FUNCTION_BLOCK TcoSequencerNonAutoRestorableTest EXTENDS TcoCore._internals_TcoContext
VAR
	_callMyPlcInstance	:	BOOL := FALSE;
	_sequencer : _TcoSequencer(THIS^, eRestoreMode.None);
	_runPLCinstanceOnce : BOOL := FALSE;
	_runPLCinstanceCyclicaly : BOOL := FALSE;
	_stepID : INT := 32764;
	_enabled : BOOL;
	_stepDescription : STRING := 'Last step sequence message';	
	_runOneStep : BOOL;
	_runAllSteps : BOOL;
	_finishStep : BOOL;
	_restore : BOOL;
	_cycleCount : INT;
	_restoreCycleCount : INT;
	_init: BOOL;
END_VAR

IF _callMyPlcInstance THEN
	IF NOT _init THEN
		ContextOpen();	
		ContextClose();	
		_init := THIS^._rtc.IsValid;
	END_IF
	
	IF _restore THEN
		ContextOpen();	
		THIS^._sequencer.Restore();	
		_restoreCycleCount := _restoreCycleCount + 1;
		_restore := FALSE;
		ContextClose();	
		RETURN;
	END_IF
	
	IF _runPLCinstanceOnce AND NOT _runPLCinstanceCyclicaly THEN
		ContextOpen();	
		THIS^.PLCinstanceRun(_stepID , _enabled, _stepDescription);
		_cycleCount := _cycleCount + 1;
		_runPLCinstanceOnce := FALSE;
		ContextClose();	
	END_IF
	
	IF _runPLCinstanceCyclicaly AND NOT _runPLCinstanceOnce THEN
		ContextOpen();	
		THIS^.PLCinstanceRun(_stepID , _enabled, _stepDescription);
		_cycleCount := _cycleCount + 1;
		ContextClose();	
	END_IF
END_IF;

{attribute 'TcRpcEnable'}
METHOD ChildHasAutoRestoreEnabled : BOOL;
ChildHasAutoRestoreEnabled := _sequencer.ChildHasAutoRestoreEnabled();
END_METHOD

{attribute 'TcRpcEnable'}
METHOD ChildIsAutoRestorable : BOOL;
ChildIsAutoRestorable := _sequencer.ChildIsAutoRestorable();
END_METHOD

{attribute 'TcRpcEnable'}
METHOD CleanupPointers
_sequencer.CleanupPointers();
END_METHOD

{attribute 'TcRpcEnable'}
METHOD ClearNumberOfSteps
_sequencer.ClearNumberOfSteps();
END_METHOD

{attribute 'TcRpcEnable'}
METHOD PROTECTED ContextClose
SUPER^._Close();
END_METHOD

{attribute 'TcRpcEnable'}
METHOD ContextOpen
SUPER^._Open();
END_METHOD

{attribute 'TcRpcEnable'}
METHOD GetChildState : INT
GetChildState := _sequencer.GetChildState();
END_METHOD

{attribute 'TcRpcEnable'}
METHOD GetCurrentStepOrder : UINT
GetCurrentStepOrder := _sequencer._currentStep.Order;
END_METHOD

{attribute 'TcRpcEnable'}
METHOD GetNumberOfStepsInSequence : UINT
GetNumberOfStepsInSequence := _sequencer._numberOfStepsInSequence;
END_METHOD

{attribute 'TcRpcEnable'}
METHOD GetOrderOfTheCurrentlyEvaluatedStep : UINT
GetOrderOfTheCurrentlyEvaluatedStep := _sequencer._theOrderOfTheCurrentlyEvaluatedStep;
END_METHOD

{attribute 'TcRpcEnable'}
METHOD GetOrderOfTheCurrentlyExecutedStep : UINT
GetOrderOfTheCurrentlyExecutedStep := _sequencer._theOrderOfTheCurrentlyExecutedStep;
END_METHOD

{attribute 'TcRpcEnable'}
METHOD GetPreviousNumberOfStepsInSequence : UINT
GetPreviousNumberOfStepsInSequence := _sequencer._previousNumberOfStepsInSequence;
END_METHOD

{attribute 'TcRpcEnable'}
METHOD GetRequestStepCycle : UINT
GetRequestStepCycle := _sequencer.RequestStepCycle;
END_METHOD

{attribute 'TcRpcEnable'}
METHOD GetSequencerErrorId : INT
GetSequencerErrorId := _sequencer.GetSequencerErrorId();
END_METHOD

{attribute 'TcRpcEnable'}
METHOD GetTextOfTheMostImportantMessage : STRING(254)
GetTextOfTheMostImportantMessage := THIS^._sequencer.GetTextOfTheMostImportantMessage();
END_METHOD

{attribute 'TcRpcEnable'}
METHOD HasAutoRestoreEnabled : BOOL;
HasAutoRestoreEnabled := _sequencer.HasAutoRestoreEnabled();
END_METHOD

{attribute 'TcRpcEnable'}
METHOD IsAutoRestorable : BOOL;
IsAutoRestorable := _sequencer.IsAutoRestorable();
END_METHOD

{attribute 'TcRpcEnable'}
METHOD IsFirstStepEntry : BOOL
IsFirstStepEntry := THIS^._sequencer.IsFirstStepEntry();
END_METHOD

METHOD PROTECTED  Main
END_METHOD

{attribute 'TcRpcEnable'}
METHOD PLCinstanceRun
VAR_INPUT
	inStepId			:	UINT;
	inEnabled			:	BOOL;
	inStepDescription	:	STRING(254);	
END_VAR
THIS^._sequencer.SetTestParams(	_runOneStep , _runAllSteps , _finishStep , inStepId , inEnabled , inStepDescription);

THIS^._sequencer.Run();
END_METHOD

{attribute 'TcRpcEnable'}
METHOD RequestStep
VAR_INPUT
	inRequestedStepId : INT;
END_VAR
_sequencer._RequestStep(inRequestedStepId);
END_METHOD

{attribute 'TcRpcEnable'}
METHOD Restore
_sequencer.Restore();
END_METHOD

{attribute 'TcRpcEnable'}
METHOD SequenceComplete
_sequencer._SequenceComplete();
END_METHOD

{attribute 'TcRpcEnable'}
METHOD SequencerClose
THIS^._sequencer.SequencerClose();
END_METHOD

{attribute 'TcRpcEnable'}
METHOD SequencerHasError : BOOL
SequencerHasError := _sequencer.SequencerHasError();
END_METHOD

{attribute 'TcRpcEnable'}
METHOD SequencerOpen
THIS^._sequencer.SequencerOpen();
END_METHOD

{attribute 'TcRpcEnable'}
METHOD SetChildState
VAR_INPUT
	inState			:	INT;
END_VAR
_sequencer.SetChildState(inState);
END_METHOD

{attribute 'TcRpcEnable'}
METHOD SetCurrentStep
VAR_INPUT
	inStepID 			:	INT;
	inStepDescription	:	STRING(254);
END_VAR
_sequencer.SetCurrentStep(inStepID := inStepID, inStepDescription := inStepDescription);
END_METHOD

{attribute 'TcRpcEnable'}
METHOD SetCurrentStepToErrorState : BOOL
SetCurrentStepToErrorState := _sequencer.SetCurrentStepToErrorState();
END_METHOD

{attribute 'TcRpcEnable'}
METHOD SetCyclicMode : BOOL
SetCyclicMode := _sequencer.SetCyclicMode();
END_METHOD

{attribute 'TcRpcEnable'}
METHOD SetInvalidMode : BOOL
SetInvalidMode := _sequencer.SetInvalidMode();
END_METHOD

{attribute 'TcRpcEnable'}
METHOD SetNumberOfSteps : UINT
VAR_INPUT
	inNumberOfSteps :UINT;
END_VAR
_sequencer.SetNumberOfSteps(inNumberOfSteps);
SetNumberOfSteps := _sequencer._numberOfStepsInSequence;
END_METHOD

{attribute 'TcRpcEnable'}
METHOD SetRequestStepCycle : UINT
VAR_INPUT
	Value : UINT;
END_VAR
_sequencer.RequestStepCycle := Value;

SetRequestStepCycle := _sequencer.RequestStepCycle;
END_METHOD

{attribute 'TcRpcEnable'}
METHOD SetSequenceAsChecked : BOOL
VAR_INPUT
END_VAR
_sequencer.SetSequenceAsChecked();
END_METHOD

{attribute 'TcRpcEnable'}
METHOD SetSequenceAsNotChecked : BOOL
VAR_INPUT
END_VAR
_sequencer.SetSequenceAsNotChecked();
END_METHOD

{attribute 'TcRpcEnable'}
METHOD SetStepMode : BOOL
SetStepMode := _sequencer.SetStepMode();
END_METHOD

{attribute 'TcRpcEnable'}
METHOD Step : BOOL
VAR_INPUT
	inStepId			:	INT;
	inEnabled			:	BOOL;
	inStepDescription	:	STRING(254);		
END_VAR
Step := _sequencer._Step(inStepID := inStepId, inEnabled := inEnabled, inStepDescription := inStepDescription);
END_METHOD

{attribute 'TcRpcEnable'}
METHOD StepBackward
_sequencer._StepBackward();
END_METHOD

{attribute 'TcRpcEnable'}
METHOD StepCompleteWhen 
VAR_INPUT
	inCondition : BOOL;
END_VAR
_sequencer._StepCompleteWhen(inCondition);
END_METHOD

{attribute 'TcRpcEnable'}
METHOD StepForward
_sequencer._StepForward();
END_METHOD

{attribute 'TcRpcEnable'}
METHOD StepIn
_sequencer._StepIn();
END_METHOD

{attribute 'TcRpcEnable'}
METHOD UpdateCurrentStepDetails
VAR_INPUT
END_VAR
_sequencer.UpdateCurrentStepDetails();
END_METHOD

END_FUNCTION_BLOCK

(* stored: Version 1.1.0.1
   POU TcoSequencerNonAutoRestorableTest: Id {8f4722b8-66cc-0a14-0d12-793c3c18c5f7}, SpecialFunc None
   Method ChildHasAutoRestoreEnabled: Id {5f6a71ef-d189-0721-3ae0-d7216f72e016}
   Method ChildIsAutoRestorable: Id {1513995a-167f-096d-2eef-38acd1e6fae4}
   Method CleanupPointers: Id {d53703e3-87a6-0d8a-1c78-693ab7549e96}
   Method ClearNumberOfSteps: Id {7f5b6809-45e4-0cee-2e5f-613b97a42248}
   Method ContextClose: Id {b958e08b-ea3d-043c-2c04-1e3f161d5009}
   Method ContextOpen: Id {79b42267-7afd-0c4f-0bbc-1b54b0e90eea}
   Method GetChildState: Id {2d71eeca-dec8-0d13-16b9-5fc527eb1f88}
   Method GetCurrentStepOrder: Id {9f0905c5-d21b-0d99-2799-a721b1fa1226}
   Method GetNumberOfStepsInSequence: Id {ece3f3c1-0aa1-01fd-3804-59fd28cfc5aa}
   Method GetOrderOfTheCurrentlyEvaluatedStep: Id {87a2cd26-1e48-002d-0d03-eaffca3cd161}
   Method GetOrderOfTheCurrentlyExecutedStep: Id {44fd8492-7e54-0a93-060d-f63030f9a407}
   Method GetPreviousNumberOfStepsInSequence: Id {089b6961-6b50-00c9-1e61-caec700a191e}
   Method GetRequestStepCycle: Id {4abdf6b0-e671-003a-3551-784d6c65cb16}
   Method GetSequencerErrorId: Id {a8e1a44f-2909-05d9-3ce0-b20390a48e05}
   Method GetTextOfTheMostImportantMessage: Id {32aafd6c-d62a-0e5d-2485-025ca9f81ee9}
   Method HasAutoRestoreEnabled: Id {b7faf085-1406-0683-07b2-6671600475aa}
   Method IsAutoRestorable: Id {adca8c3f-c81e-0f3c-311d-8e51e07b5c8a}
   Method IsFirstStepEntry: Id {a7030725-a7ca-088c-35b1-f3dce620f31e}
   Method Main: Id {42cb7ad9-ea6a-0869-1918-2e4efedffd1d}
   Method PLCinstanceRun: Id {284fbd9f-5e0b-066a-3e75-1b2389860cb3}
   Method RequestStep: Id {e9a05251-1aa2-09a6-1293-ede5ed4234e5}
   Method Restore: Id {1ef21be0-22b9-0ca7-080d-885fdb40798f}
   Method SequenceComplete: Id {3a8cf623-e5e1-0266-2042-a382cbeb5fd5}
   Method SequencerClose: Id {2db8b4a8-0cb6-0018-3fd0-1a932fae0a02}
   Method SequencerHasError: Id {d27f0ba1-15ec-0fff-027b-579d89ee6265}
   Method SequencerOpen: Id {9b07bafb-4d05-0518-0fa5-898b5160b2bf}
   Method SetChildState: Id {12342cf7-42b9-03d2-1c7f-3794e8186cb8}
   Method SetCurrentStep: Id {d2f7209a-4095-09a1-156f-bb1bb625d606}
   Method SetCurrentStepToErrorState: Id {62518721-0247-0b6c-2e49-d0dd0f36718c}
   Method SetCyclicMode: Id {d0feb316-77b3-0136-1521-af6499a4203a}
   Method SetInvalidMode: Id {a9a29389-049b-02f7-2034-6345e249d17a}
   Method SetNumberOfSteps: Id {4327b4be-d6a7-0f65-2cf9-4478d1a488e5}
   Method SetRequestStepCycle: Id {eaba7156-f498-0d8b-357d-f086640e0b79}
   Method SetSequenceAsChecked: Id {3875aa8f-d84f-0c02-31a6-cacbc68b8826}
   Method SetSequenceAsNotChecked: Id {20c162cf-155b-068f-2e24-fa0c35deb5fd}
   Method SetStepMode: Id {323a566b-5dc2-0b7f-1e3c-83dc699013ca}
   Method Step: Id {efa0cec6-6d10-0a3d-286c-9b1e1dd7f678}
   Method StepBackward: Id {4186a26f-6755-0eb7-3e54-bdaf5b8b4f1a}
   Method StepCompleteWhen: Id {b3705be5-f91d-0220-0744-1d62aceb9806}
   Method StepForward: Id {64ba9f52-e7ce-019a-16db-ac9127859354}
   Method StepIn: Id {51e40032-50ea-050e-279a-323a8bbf0a82}
   Method UpdateCurrentStepDetails: Id {704b1d04-ff8c-0f27-1c43-63c0df064c73} *)
